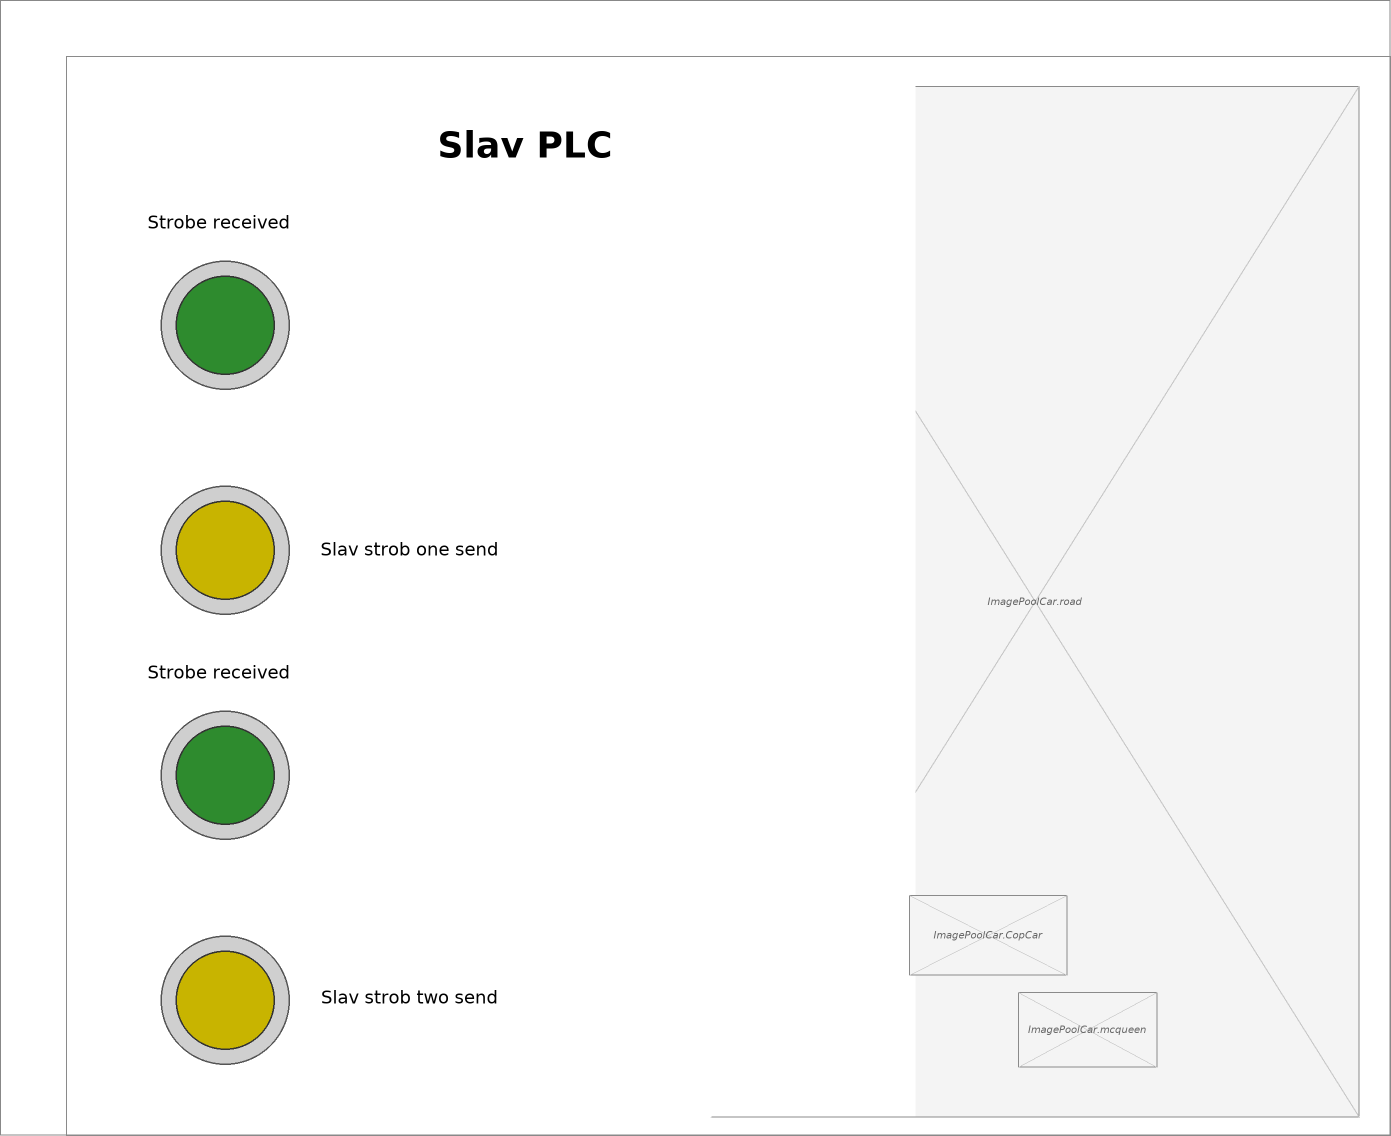
VISUALIZATION VisualizationSlave  // 1391x1136
    Frame (66,56 1325x1080)
    Image (711,86 648x1031), image: ImagePoolCar.road
    Rectangle (637,86 278x1030)
    Label (400,120 250x50), "Slav PLC"
    Lamp1 (150,250 150x150), variable: GVLSlave.OXLampIXOneGreen, style: Lamp-Lamp1-Green
    Label (100,200 238x45), "Strobe received"
    Label (300,527 219x45), "Slav strob one send"
    Lamp1 (150,475 150x150), variable: GVLSlave.OXLampOXOne, style: Lamp-Lamp1-Yellow
    Lamp1 (150,700 150x150), variable: GVLSlave.OXLampIXTwoGreen, style: Lamp-Lamp1-Green
    Lamp1 (150,925 150x150), variable: GVLSlave.OXLampOXTwo, style: Lamp-Lamp1-Yellow
    Image (1018,992 139x75), angle 90, image: ImagePoolCar.mcqueen
        p3528305787: GVLSlave.OIntRedCar
        p874137650: GVLSlave.OIntRedCar
    Image (909,895 158x80), angle 90, image: ImagePoolCar.CopCar
        p3528305787: GVLSlave.OintCopCar
        p874137650: GVLSlave.OintCopCar
    Label (300,975 219x45), "Slav strob two send"
    Label (100,650 238x45), "Strobe received"
    Label (450,650 150x30)
END_VISUALIZATION

(* stored: Version 1.1.0.1, ProductVersion 3.1.4024.12
   Visu VisualizationSlave: Id {77b04896-c5a4-43e9-805c-d96302aa5f75} *)
